Staubli VAL3: switchItem.pjx

--- switchItem.pjx ---
Parameters version=s8.12.1Cs9_BS2449 stackSize=5000 millimeterUnit=true
Data file=switchItem.dtx

--- switchItem.dtx ---
public num nSwitchValue
public string sIOValue
public bool bIOdisable
